(* IEC 61131-3 sources: model-first-plc-agent-ai/results/T2-W-24, 2 files *)

(* ---- a1_code.st ---- *)
FUNCTION_BLOCK TankRuntime
VAR_INPUT
    start : BOOL;
    stop : BOOL;
    LSH : BOOL;
    LSHH : BOOL;
    TimerDuration : TIME;
END_VAR
VAR_OUTPUT
    fill_valve : BOOL;
    discharge_valve : BOOL;
END_VAR
VAR
    x0 : BOOL := TRUE;
    x1 : BOOL := FALSE;
    timer_done : BOOL := FALSE;
    FillingTimer : TON;
    transition_start : BOOL;
    transition_finish : BOOL;
END_VAR

(* Evaluate the timer for the currently active situation. *)
FillingTimer(IN := x1, PT := TimerDuration);
timer_done := FillingTimer.Q;

(* Evaluate both transitions before changing the active situation. *)
transition_start := x0 AND start AND NOT stop AND NOT LSHH;
transition_finish := x1 AND (stop OR LSHH OR timer_done);

IF transition_finish THEN
    x0 := TRUE;
    x1 := FALSE;

    (* Reset the owned timer immediately on leaving x1. *)
    FillingTimer(IN := FALSE, PT := TimerDuration);
    timer_done := FALSE;

ELSIF transition_start THEN
    x0 := FALSE;
    x1 := TRUE;

    (* Start timing immediately on entering x1. *)
    FillingTimer(IN := TRUE, PT := TimerDuration);
    timer_done := FALSE;
END_IF;

fill_valve := x1;
discharge_valve := FALSE;

END_FUNCTION_BLOCK

PROGRAM Main
VAR
    StartCommand AT %IX100.0 : BOOL;
    StopCommand AT %IX100.1 : BOOL;
    LSH AT %IX100.2 : BOOL;
    LSHH AT %IX100.3 : BOOL;
    FillValve AT %QX100.0 : BOOL;
    DischargeValve AT %QX100.1 : BOOL;
END_VAR
VAR
    (* Configurable filling interval. *)
    TimerDuration : TIME := T#10s;
    StartEdge : R_TRIG;
    TankControl : TankRuntime;
END_VAR

StartEdge(CLK := StartCommand);

TankControl(
    start := StartEdge.Q,
    stop := StopCommand,
    LSH := LSH,
    LSHH := LSHH,
    TimerDuration := TimerDuration
);

FillValve := TankControl.fill_valve;
DischargeValve := TankControl.discharge_valve;

END_PROGRAM

(* ---- a2_code.st ---- *)
FUNCTION_BLOCK FB_TimedTankFilling
VAR_INPUT
    StartCommand : BOOL;
    StopCommand : BOOL;
    LSH : BOOL;
    LSHH : BOOL;
    TimerDuration : TIME;
END_VAR
VAR_OUTPUT
    fill_valve : BOOL;
    discharge_valve : BOOL;
END_VAR
VAR
    StartEdge : R_TRIG;
    FillingTimer : TON;
    start : BOOL;
    stop : BOOL;
    timer_done : BOOL;
    FillingState : INT := 0;
END_VAR

StartEdge(CLK := StartCommand);
start := StartEdge.Q;
stop := StopCommand;

IF stop THEN
    FillingState := 0;
ELSIF FillingState = 0 THEN
    IF start AND NOT LSHH THEN
        FillingState := 1;
    END_IF;
ELSIF FillingState <> 1 THEN
    FillingState := 0;
END_IF;

(* Timing begins in the scan that activates the filling step. *)
FillingTimer(
    IN := (FillingState = 1),
    PT := TimerDuration
);
timer_done := FillingTimer.Q;

IF FillingState = 1 THEN
    IF stop OR LSHH OR timer_done THEN
        FillingState := 0;

        (* Reset the step-owned timer immediately upon leaving filling. *)
        FillingTimer(IN := FALSE, PT := TimerDuration);
        timer_done := FillingTimer.Q;
    END_IF;
END_IF;

fill_valve := (FillingState = 1);
discharge_valve := FALSE;

END_FUNCTION_BLOCK

PROGRAM Main
VAR
    StartCommand AT %IX100.0 : BOOL;
    StopCommand AT %IX100.1 : BOOL;
    LSH AT %IX100.2 : BOOL;
    LSHH AT %IX100.3 : BOOL;
    FillValve AT %QX100.0 : BOOL;
    DischargeValve AT %QX100.1 : BOOL;
END_VAR
VAR
    TankController : FB_TimedTankFilling;
    TimerDuration : TIME := T#10s; (* Configurable filling-time preset. *)
END_VAR

TankController(
    StartCommand := StartCommand,
    StopCommand := StopCommand,
    LSH := LSH,
    LSHH := LSHH,
    TimerDuration := TimerDuration
);

FillValve := TankController.fill_valve;
DischargeValve := TankController.discharge_valve;

END_PROGRAM
